// SIMATIC S7-200 project (STEP 7-Micro/WIN), CPU 224XP CN REL 02.01

ORGANIZATION_BLOCK PRINCIPAL:OB1
TITLE=COMENTARIOS DEL PROGRAMA
BEGIN
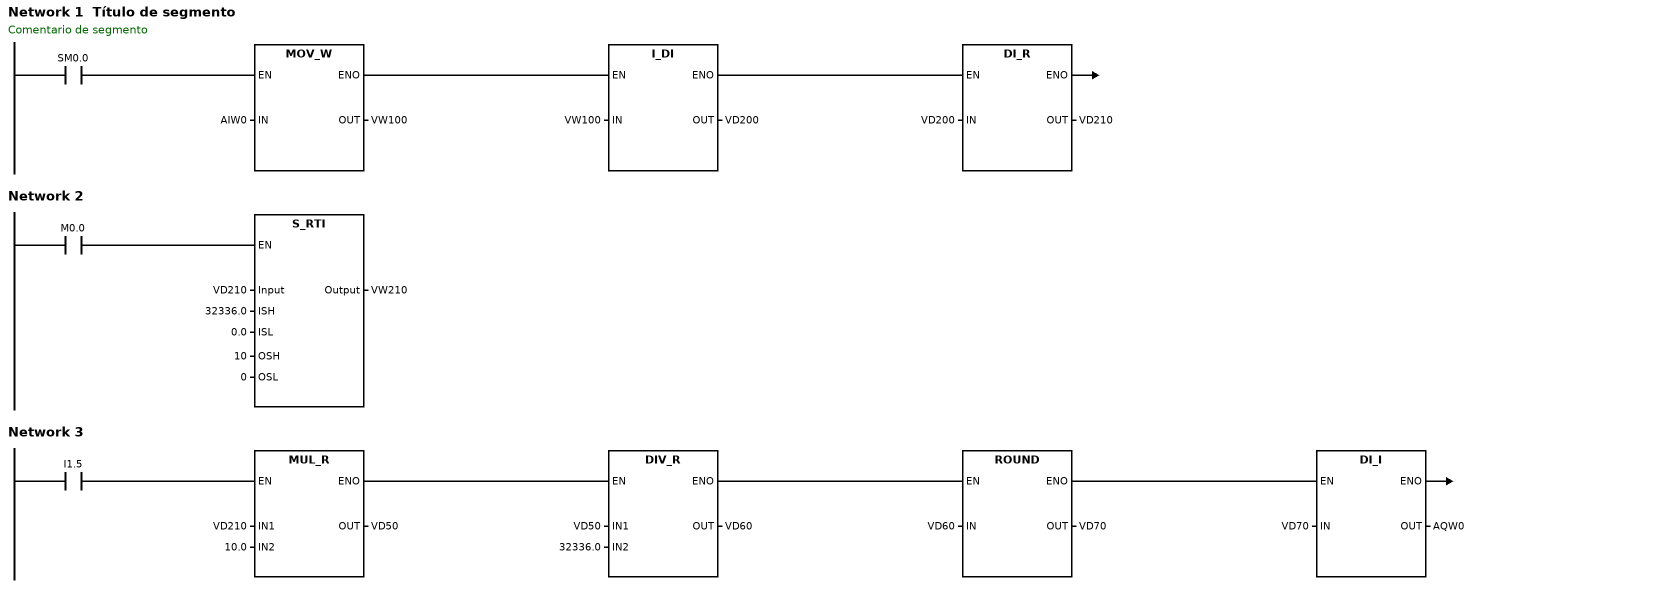
Network 1 // Título de segmento
// Comentario de segmento
LD     SM0.0
MOVW   AIW0, VW100
AENO
ITD    VW100, VD200
AENO
DTR    VD200, VD210
Network 2
LD     M0.0
CALL   S_RTI:SBR1, VD210, 32336.0, 0.0, 10, 0, VW210
Network 3
LD     I1.5
MOVR   VD210, VD50
AENO
*R     10.0, VD50
AENO
MOVR   VD50, VD60
AENO
/R     32336.0, VD60
AENO
ROUND  VD60, VD70
AENO
DTI    VD70, AQW0
END_ORGANIZATION_BLOCK

// SBR1: protected block, not included
